Staubli VAL3: init.pgx

public program init()
  local num l_i
begin
  nPage=0
  nPageIndex=0
  nItemIndex=0

  nPage=roundUp(size(io:dInItem)/16)
  sShowPageIndex=toString("",nPageIndex+1)
  sPageNum=toString("",nPage)
  sUsingBus=rs:sBusUsing
  nSelType=0
  call SetbtnColor(nSelType)
  for l_i = 0 to 15
    sLabel[l_i]=""
    sComment[l_i]=""
  endFor
  if io:nMaxAnalog<=0
    userPageSet("IO","btn3","disabled",true)
    userPageSet("IO","btn4","disabled",true)
    popUpMsg("模拟量数量未设置")
  endIf
  //  //list
  //  for l_i = 0 to 15
  //    sLabel[l_i]="dIn["+toString("",l_i+16*nPageIndex)+"]"
  //    sComment[l_i]=io:dInItem[l_i+16*nPageIndex].sComment
  //  endFor

end
